Fanuc KAREL source: kb00202.KL

-- PROVISIONAL review KL for V1013-1; original PC SHA256 39569739d6a6c9f8f5ba7818886c6618e79802f7d0eb12f3192798954f5f8598
-- Incomplete behavior may be omitted. Consult companion uncertainty JSON. Do not deploy.
PROGRAM KB00202
%NOLOCKGROUP
BEGIN
  -- UNRESOLVED_PC offsets 5-14; opcodes 3F,75
  -- UNRESOLVED_PC offsets 19-28; opcodes 3F,75
  -- UNRESOLVED_PC offsets 33-40; opcodes 9D,23
  -- UNRESOLVED_PC offsets 45-77; opcodes 27,22,22,2A,22,2A,22,31
  -- UNRESOLVED_PC offsets 82-86; opcodes 7F
END KB00202
